(* IEC 61131-3 sources: POMIRTS_lab3/AS/Library_2/AsICMP, 3 files *)

(* ---- AsICMP.typ ---- *)
TYPE

END_TYPE

(* ---- AsICMP.fun ---- *)
{REDUND_CONTEXT} {REDUND_UNREPLICABLE} FUNCTION_BLOCK IcmpPing					(*pings a station; asynchronous execution*)
	VAR_INPUT
		enable			: BOOL;			(*enables execution*)
		pHost			: UDINT;		(*pointer to the IP address or name of the station that should be pinged*)
		timeout			: UINT;			(*response timeout*)
	END_VAR

	VAR_OUTPUT
		status			: UINT;			(*execution status: ERR_OK, ERR_FUB_ENABLE_FALSE, ERR_FUB_BUSY, 0xXXXX = see help*)
	END_VAR

	VAR
        i_state			: UINT;			(*internal variable*)
		i_result		: UINT;			(*internal variable*)
        i_tmp			: UDINT;		(*internal variable*)
	END_VAR
END_FUNCTION_BLOCK

(* ---- AsICMP.var ---- *)
VAR CONSTANT
	icmpERR_NO_RESPONSE					: UINT := 32750;	(*no ping response*)
	icmpERR_PARAMETER					: UINT := 32751;	(*invalid parameter, check parameter*)
	icmpERR_SOCKET_CREATE				: UINT := 32752;	(*create socket failed*)
	icmpERR_UNREACHABLE					: UINT := 32753;	(*host unreachable*)
	icmpERR_SYSTEM						: UINT := 32799;	(*system error*)
END_VAR
